// LS Electric XG5000 project: 1조_2차_2축_공압+로드셀_최종
// PLC LSPLC
// module base 0 slot 0: Input/Output Module:XBM-DN/DP32H2 (DC 24V Input/TR Output, 32 points)
// module base 0 slot 1: Internal Positioning:XBF-PO02E (Open Collector Type, 2 Axis)
// module base 0 slot 2: Positioning Module:XBF-PN04B (Position Control, EtherCAT Network Type(4 axis))
// module base 0 slot 3: Loadcell Input Module:XBF-LD02S (Isolated-type Loadcell Input(2 Channels))
// task INIT: Kind=1 Priority=2

PROGRAM ERROR (task: 스캔 프로그램)

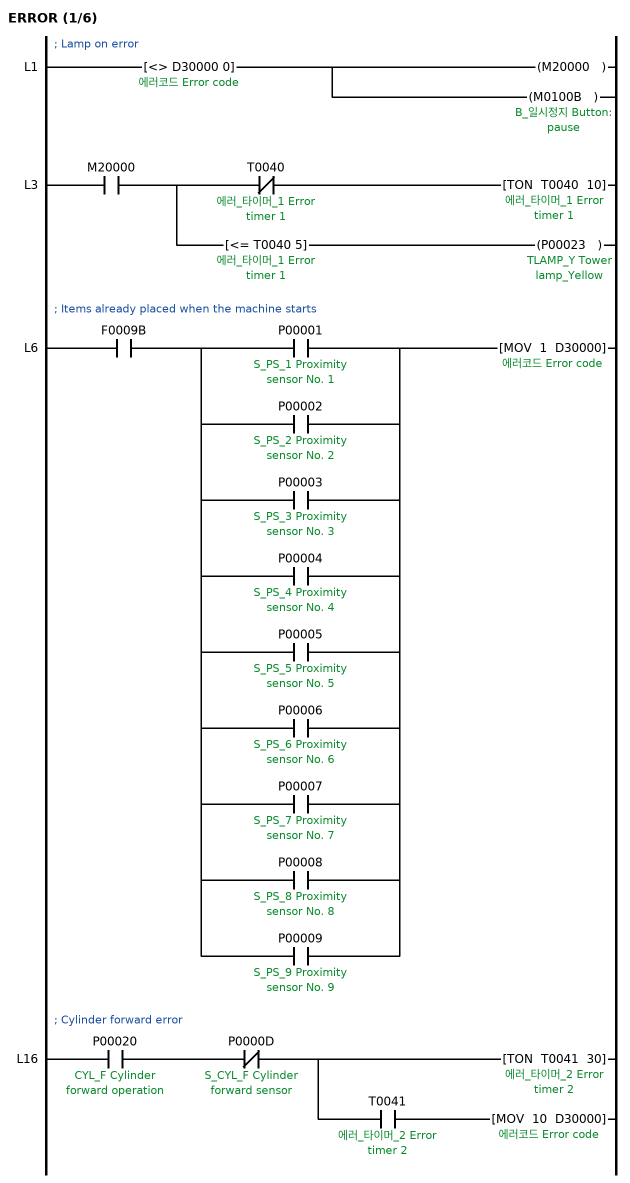
// Lamp on error
; L1
LOAD<>    D30000 0	// 에러코드 Error code
OUT       M20000
OUT       M0100B	// B_일시정지 Button: pause
; L3
LOAD      M20000
MPUSH
AND NOT   T0040	// 에러_타이머_1 Error timer 1
TON       T0040 10	// 에러_타이머_1 Error timer 1
MPOP
AND<=     T0040 5	// 에러_타이머_1 Error timer 1
OUT       P00023	// TLAMP_Y Tower lamp_Yellow
// Items already placed when the machine starts
; L6
LOAD      F0009B
LOAD      P00001	// S_PS_1 Proximity sensor No. 1
OR        P00002	// S_PS_2 Proximity sensor No. 2
OR        P00003	// S_PS_3 Proximity sensor No. 3
OR        P00004	// S_PS_4 Proximity sensor No. 4
OR        P00005	// S_PS_5 Proximity sensor No. 5
OR        P00006	// S_PS_6 Proximity sensor No. 6
OR        P00007	// S_PS_7 Proximity sensor No. 7
OR        P00008	// S_PS_8 Proximity sensor No. 8
OR        P00009	// S_PS_9 Proximity sensor No. 9
AND LOAD
MOV       1 D30000	// 에러코드 Error code
// Cylinder forward error
; L16
LOAD      P00020	// CYL_F Cylinder forward operation
AND NOT   P0000D	// S_CYL_F Cylinder forward sensor
TON       T0041 30	// 에러_타이머_2 Error timer 2
AND       T0041	// 에러_타이머_2 Error timer 2
MOV       10 D30000	// 에러코드 Error code

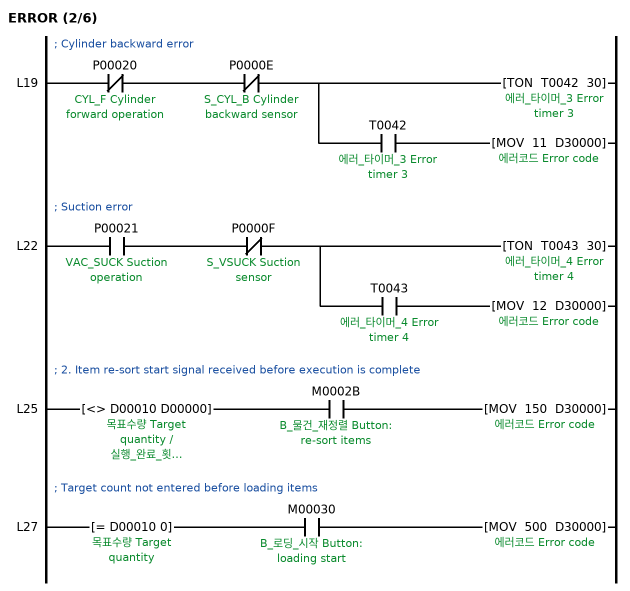
// Cylinder backward error
; L19
LOAD NOT  P00020	// CYL_F Cylinder forward operation
AND NOT   P0000E	// S_CYL_B Cylinder backward sensor
TON       T0042 30	// 에러_타이머_3 Error timer 3
AND       T0042	// 에러_타이머_3 Error timer 3
MOV       11 D30000	// 에러코드 Error code
// Suction error
; L22
LOAD      P00021	// VAC_SUCK Suction operation
AND NOT   P0000F	// S_VSUCK Suction sensor
TON       T0043 30	// 에러_타이머_4 Error timer 4
AND       T0043	// 에러_타이머_4 Error timer 4
MOV       12 D30000	// 에러코드 Error code
// 2. Item re-sort start signal received before execution is complete
; L25
LOAD<>    D00010 D00000	// 목표수량 Target quantity / 실행_완료_횟수 Execution complete count
AND       M0002B	// B_물건_재정렬 Button: re-sort items
MOV       150 D30000	// 에러코드 Error code
// Target count not entered before loading items
; L27
LOAD=     D00010 0	// 목표수량 Target quantity
AND       M00030	// B_로딩_시작 Button: loading start
MOV       500 D30000	// 에러코드 Error code

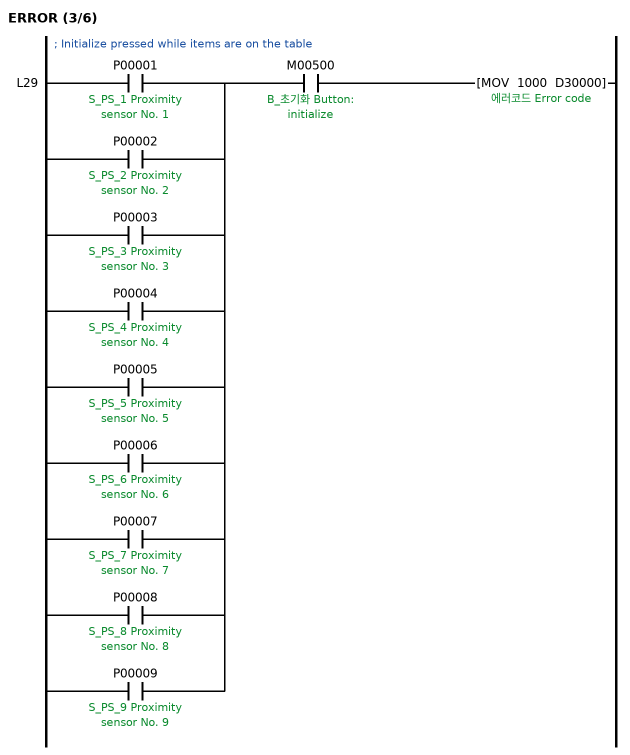
// Initialize pressed while items are on the table
; L29
LOAD      P00001	// S_PS_1 Proximity sensor No. 1
OR        P00002	// S_PS_2 Proximity sensor No. 2
OR        P00003	// S_PS_3 Proximity sensor No. 3
OR        P00004	// S_PS_4 Proximity sensor No. 4
OR        P00005	// S_PS_5 Proximity sensor No. 5
OR        P00006	// S_PS_6 Proximity sensor No. 6
OR        P00007	// S_PS_7 Proximity sensor No. 7
OR        P00008	// S_PS_8 Proximity sensor No. 8
OR        P00009	// S_PS_9 Proximity sensor No. 9
AND       M00500	// B_초기화 Button: initialize
MOV       1000 D30000	// 에러코드 Error code

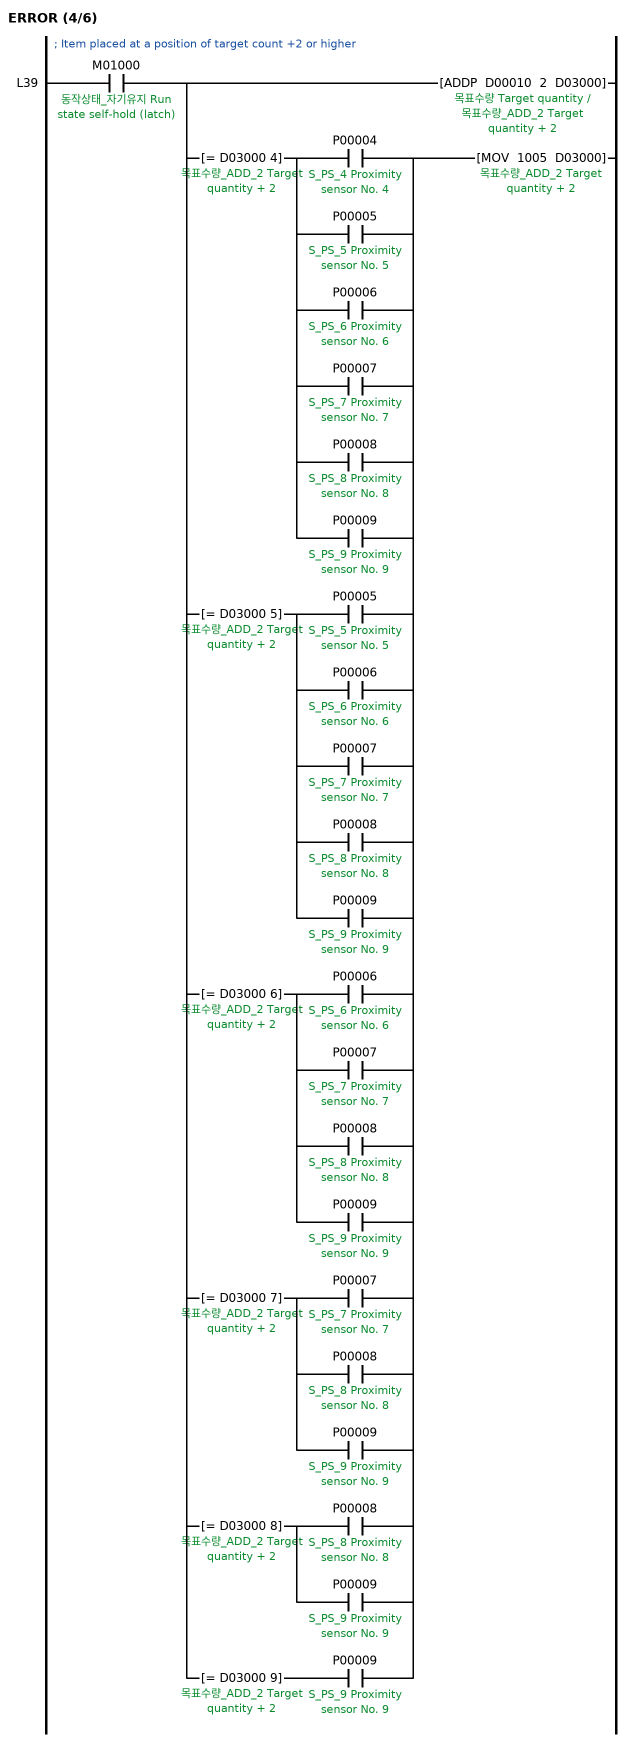
// Item placed at a position of target count +2 or higher
; L39
LOAD      M01000	// 동작상태_자기유지 Run state self-hold (latch)
ADDP      D00010 2 D03000	// 목표수량 Target quantity / 목표수량_ADD_2 Target quantity + 2
LOAD=     D03000 4	// 목표수량_ADD_2 Target quantity + 2
LOAD      P00004	// S_PS_4 Proximity sensor No. 4
OR        P00005	// S_PS_5 Proximity sensor No. 5
OR        P00006	// S_PS_6 Proximity sensor No. 6
OR        P00007	// S_PS_7 Proximity sensor No. 7
OR        P00008	// S_PS_8 Proximity sensor No. 8
OR        P00009	// S_PS_9 Proximity sensor No. 9
AND LOAD
LOAD=     D03000 5	// 목표수량_ADD_2 Target quantity + 2
LOAD      P00005	// S_PS_5 Proximity sensor No. 5
OR        P00006	// S_PS_6 Proximity sensor No. 6
OR        P00007	// S_PS_7 Proximity sensor No. 7
OR        P00008	// S_PS_8 Proximity sensor No. 8
OR        P00009	// S_PS_9 Proximity sensor No. 9
AND LOAD
OR LOAD
LOAD=     D03000 6	// 목표수량_ADD_2 Target quantity + 2
LOAD      P00006	// S_PS_6 Proximity sensor No. 6
OR        P00007	// S_PS_7 Proximity sensor No. 7
OR        P00008	// S_PS_8 Proximity sensor No. 8
OR        P00009	// S_PS_9 Proximity sensor No. 9
AND LOAD
OR LOAD
LOAD=     D03000 7	// 목표수량_ADD_2 Target quantity + 2
LOAD      P00007	// S_PS_7 Proximity sensor No. 7
OR        P00008	// S_PS_8 Proximity sensor No. 8
OR        P00009	// S_PS_9 Proximity sensor No. 9
AND LOAD
OR LOAD
LOAD=     D03000 8	// 목표수량_ADD_2 Target quantity + 2
LOAD      P00008	// S_PS_8 Proximity sensor No. 8
OR        P00009	// S_PS_9 Proximity sensor No. 9
AND LOAD
OR LOAD
LOAD=     D03000 9	// 목표수량_ADD_2 Target quantity + 2
AND       P00009	// S_PS_9 Proximity sensor No. 9
OR LOAD
AND LOAD
MOV       1005 D03000	// 목표수량_ADD_2 Target quantity + 2

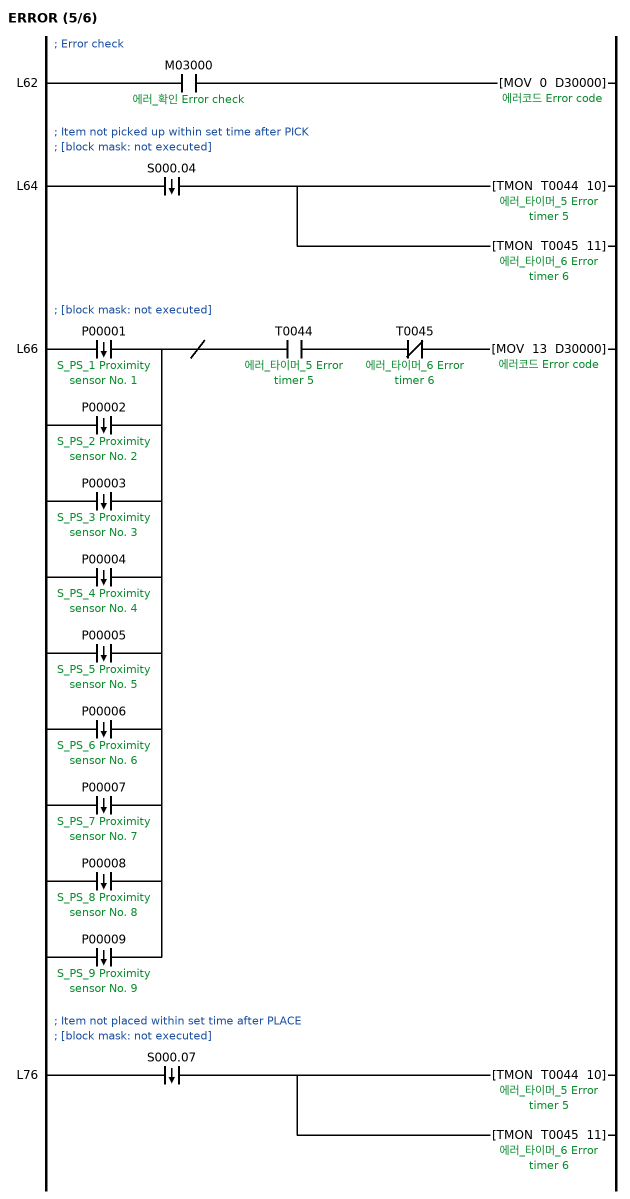
// Error check
; L62
LOAD      M03000	// 에러_확인 Error check
MOV       0 D30000	// 에러코드 Error code
// Item not picked up within set time after PICK
; L64 (block mask: not executed)
LOADN     S000.04
TMON      T0044 10	// 에러_타이머_5 Error timer 5
TMON      T0045 11	// 에러_타이머_6 Error timer 6
; L66 (block mask: not executed)
LOADN     P00001	// S_PS_1 Proximity sensor No. 1
ORN       P00002	// S_PS_2 Proximity sensor No. 2
ORN       P00003	// S_PS_3 Proximity sensor No. 3
ORN       P00004	// S_PS_4 Proximity sensor No. 4
ORN       P00005	// S_PS_5 Proximity sensor No. 5
ORN       P00006	// S_PS_6 Proximity sensor No. 6
ORN       P00007	// S_PS_7 Proximity sensor No. 7
ORN       P00008	// S_PS_8 Proximity sensor No. 8
ORN       P00009	// S_PS_9 Proximity sensor No. 9
NOT
AND       T0044	// 에러_타이머_5 Error timer 5
AND NOT   T0045	// 에러_타이머_6 Error timer 6
MOV       13 D30000	// 에러코드 Error code
// Item not placed within set time after PLACE
; L76 (block mask: not executed)
LOADN     S000.07
TMON      T0044 10	// 에러_타이머_5 Error timer 5
TMON      T0045 11	// 에러_타이머_6 Error timer 6

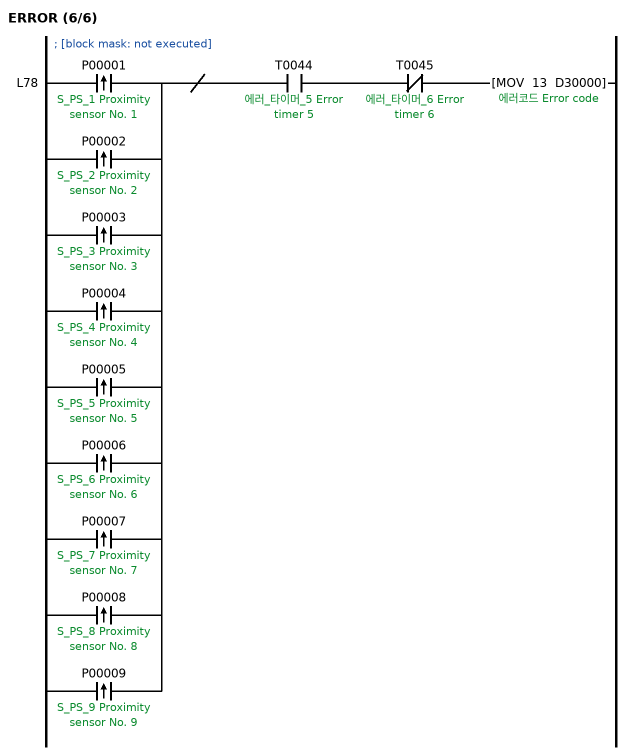
; L78 (block mask: not executed)
LOADP     P00001	// S_PS_1 Proximity sensor No. 1
ORP       P00002	// S_PS_2 Proximity sensor No. 2
ORP       P00003	// S_PS_3 Proximity sensor No. 3
ORP       P00004	// S_PS_4 Proximity sensor No. 4
ORP       P00005	// S_PS_5 Proximity sensor No. 5
ORP       P00006	// S_PS_6 Proximity sensor No. 6
ORP       P00007	// S_PS_7 Proximity sensor No. 7
ORP       P00008	// S_PS_8 Proximity sensor No. 8
ORP       P00009	// S_PS_9 Proximity sensor No. 9
NOT
AND       T0044	// 에러_타이머_5 Error timer 5
AND NOT   T0045	// 에러_타이머_6 Error timer 6
MOV       13 D30000	// 에러코드 Error code

PROGRAM Servo (task: 스캔 프로그램)

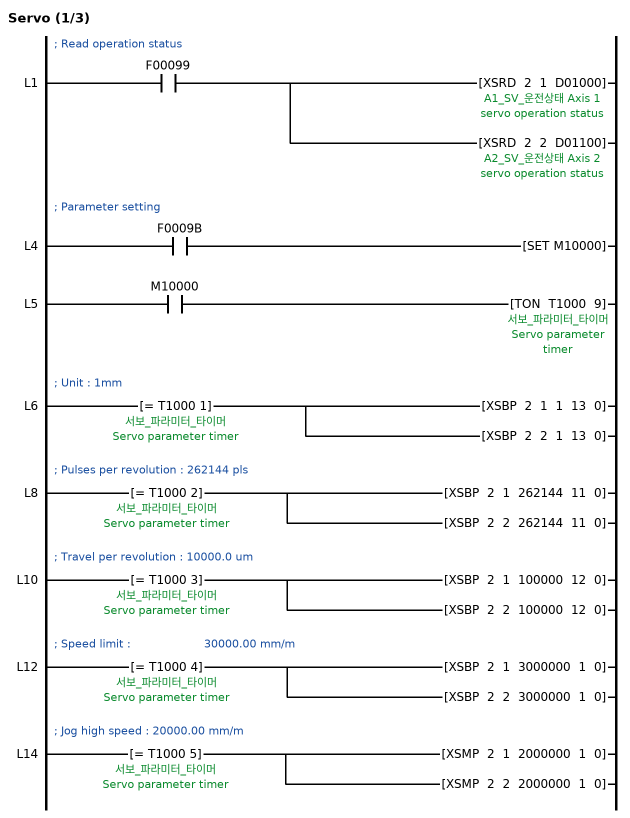
// Read operation status
; L1
LOAD      F00099
XSRD      2 1 D01000	// A1_SV_운전상태 Axis 1 servo operation status
XSRD      2 2 D01100	// A2_SV_운전상태 Axis 2 servo operation status
// Parameter setting
; L4
LOAD      F0009B
SET       M10000
; L5
LOAD      M10000
TON       T1000 9	// 서보_파라미터_타이머 Servo parameter timer
; L6
LOAD=     T1000 1	// 서보_파라미터_타이머 Servo parameter timer
XSBP      2 1 1 13 0
XSBP      2 2 1 13 0
// output comment: Unit : 1mm
; L8
LOAD=     T1000 2	// 서보_파라미터_타이머 Servo parameter timer
XSBP      2 1 262144 11 0
XSBP      2 2 262144 11 0
// output comment: Pulses per revolution : 262144 pls
; L10
LOAD=     T1000 3	// 서보_파라미터_타이머 Servo parameter timer
XSBP      2 1 100000 12 0
XSBP      2 2 100000 12 0
// output comment: Travel per revolution : 10000.0 um
; L12
LOAD=     T1000 4	// 서보_파라미터_타이머 Servo parameter timer
XSBP      2 1 3000000 1 0
XSBP      2 2 3000000 1 0
// output comment: Speed limit :                     30000.00 mm/m
; L14
LOAD=     T1000 5	// 서보_파라미터_타이머 Servo parameter timer
XSMP      2 1 2000000 1 0
XSMP      2 2 2000000 1 0
// output comment: Jog high speed : 20000.00 mm/m

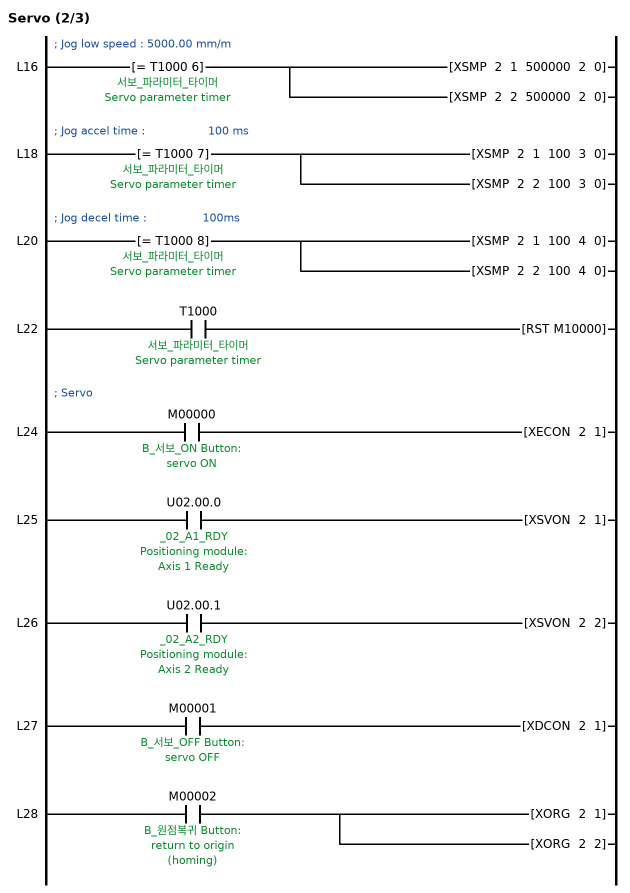
; L16
LOAD=     T1000 6	// 서보_파라미터_타이머 Servo parameter timer
XSMP      2 1 500000 2 0
XSMP      2 2 500000 2 0
// output comment: Jog low speed : 5000.00 mm/m
; L18
LOAD=     T1000 7	// 서보_파라미터_타이머 Servo parameter timer
XSMP      2 1 100 3 0
XSMP      2 2 100 3 0
// output comment: Jog accel time :                  100 ms
; L20
LOAD=     T1000 8	// 서보_파라미터_타이머 Servo parameter timer
XSMP      2 1 100 4 0
XSMP      2 2 100 4 0
// output comment: Jog decel time :                100ms
; L22
LOAD      T1000	// 서보_파라미터_타이머 Servo parameter timer
RST       M10000
// Servo
; L24
LOAD      M00000	// B_서보_ON Button: servo ON
XECON     2 1
; L25
LOAD      U02.00.0	// _02_A1_RDY Positioning module: Axis 1 Ready
XSVON     2 1
; L26
LOAD      U02.00.1	// _02_A2_RDY Positioning module: Axis 2 Ready
XSVON     2 2
; L27
LOAD      M00001	// B_서보_OFF Button: servo OFF
XDCON     2 1
; L28
LOAD      M00002	// B_원점복귀 Button: return to origin (homing)
XORG      2 1
XORG      2 2

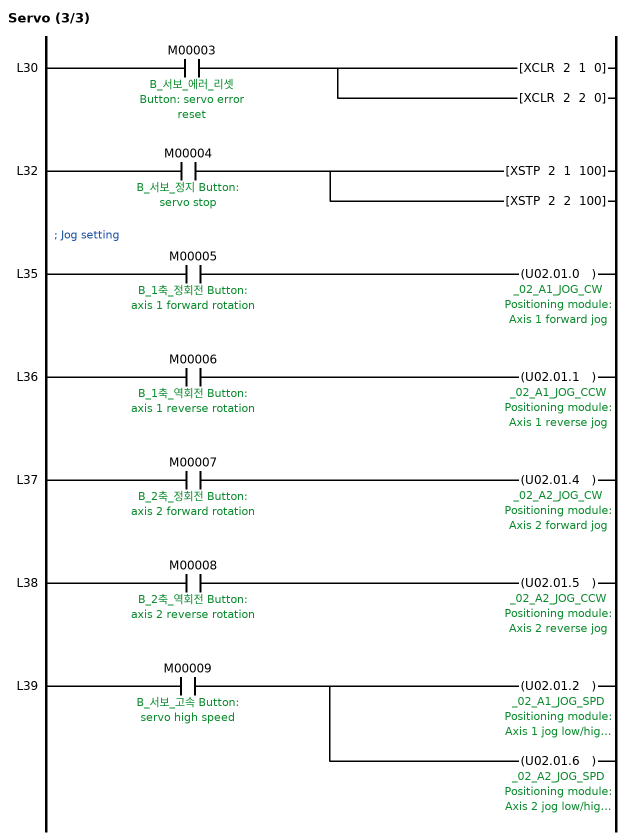
; L30
LOAD      M00003	// B_서보_에러_리셋 Button: servo error reset
XCLR      2 1 0
XCLR      2 2 0
; L32
LOAD      M00004	// B_서보_정지 Button: servo stop
XSTP      2 1 100
XSTP      2 2 100
// Jog setting
; L35
LOAD      M00005	// B_1축_정회전 Button: axis 1 forward rotation
OUT       U02.01.0	// _02_A1_JOG_CW Positioning module: Axis 1 forward jog
; L36
LOAD      M00006	// B_1축_역회전 Button: axis 1 reverse rotation
OUT       U02.01.1	// _02_A1_JOG_CCW Positioning module: Axis 1 reverse jog
; L37
LOAD      M00007	// B_2축_정회전 Button: axis 2 forward rotation
OUT       U02.01.4	// _02_A2_JOG_CW Positioning module: Axis 2 forward jog
; L38
LOAD      M00008	// B_2축_역회전 Button: axis 2 reverse rotation
OUT       U02.01.5	// _02_A2_JOG_CCW Positioning module: Axis 2 reverse jog
; L39
LOAD      M00009	// B_서보_고속 Button: servo high speed
OUT       U02.01.2	// _02_A1_JOG_SPD Positioning module: Axis 1 jog low/high speed
OUT       U02.01.6	// _02_A2_JOG_SPD Positioning module: Axis 2 jog low/high speed

PROGRAM Load_Cell (task: 스캔 프로그램)

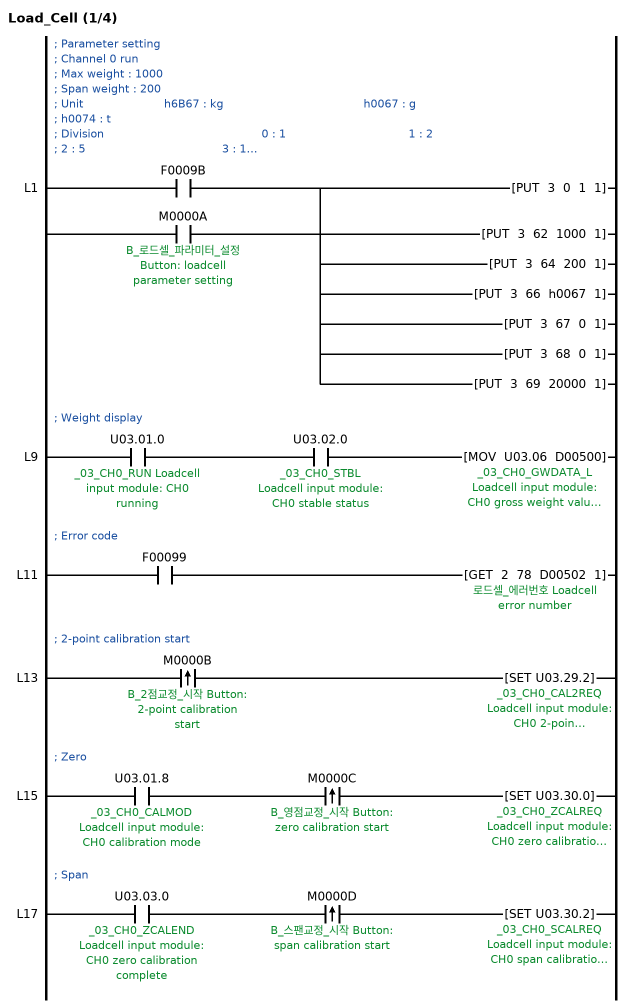
// Parameter setting
; L1
LOAD      F0009B
OR        M0000A	// B_로드셀_파라미터_설정 Button: loadcell parameter setting
PUT       3 0 1 1
PUT       3 62 1000 1
PUT       3 64 200 1
PUT       3 66 h0067 1
PUT       3 67 0 1
PUT       3 68 0 1
PUT       3 69 20000 1
// output comment: Channel 0 run
// output comment: Max weight : 1000
// output comment: Span weight : 200
// output comment: Unit                       h6B67 : kg                                        h0067 : g                                         h0074 : t
// output comment: Division                                             0 : 1                                   1 : 2                                             2 : 5                                       3 : 10
// output comment: Decimal                    0 : 1                    1: 0.1                         2 : 0.01                  3 : 0.001
// output comment: Loadcell sensitivity : 2mV/V
// Weight display
; L9
LOAD      U03.01.0	// _03_CH0_RUN Loadcell input module: CH0 running
AND       U03.02.0	// _03_CH0_STBL Loadcell input module: CH0 stable status
MOV       U03.06 D00500	// _03_CH0_GWDATA_L Loadcell input module: CH0 gross weight value (low) / Mass
// Error code
; L11
LOAD      F00099
GET       2 78 D00502 1	// 로드셀_에러번호 Loadcell error number
// 2-point calibration start
; L13
LOADP     M0000B	// B_2점교정_시작 Button: 2-point calibration start
SET       U03.29.2	// _03_CH0_CAL2REQ Loadcell input module: CH0 2-point calibration mode request
// Zero
; L15
LOAD      U03.01.8	// _03_CH0_CALMOD Loadcell input module: CH0 calibration mode
ANDP      M0000C	// B_영점교정_시작 Button: zero calibration start
SET       U03.30.0	// _03_CH0_ZCALREQ Loadcell input module: CH0 zero calibration command
// Span
; L17
LOAD      U03.03.0	// _03_CH0_ZCALEND Loadcell input module: CH0 zero calibration complete
ANDP      M0000D	// B_스팬교정_시작 Button: span calibration start
SET       U03.30.2	// _03_CH0_SCALREQ Loadcell input module: CH0 span calibration command

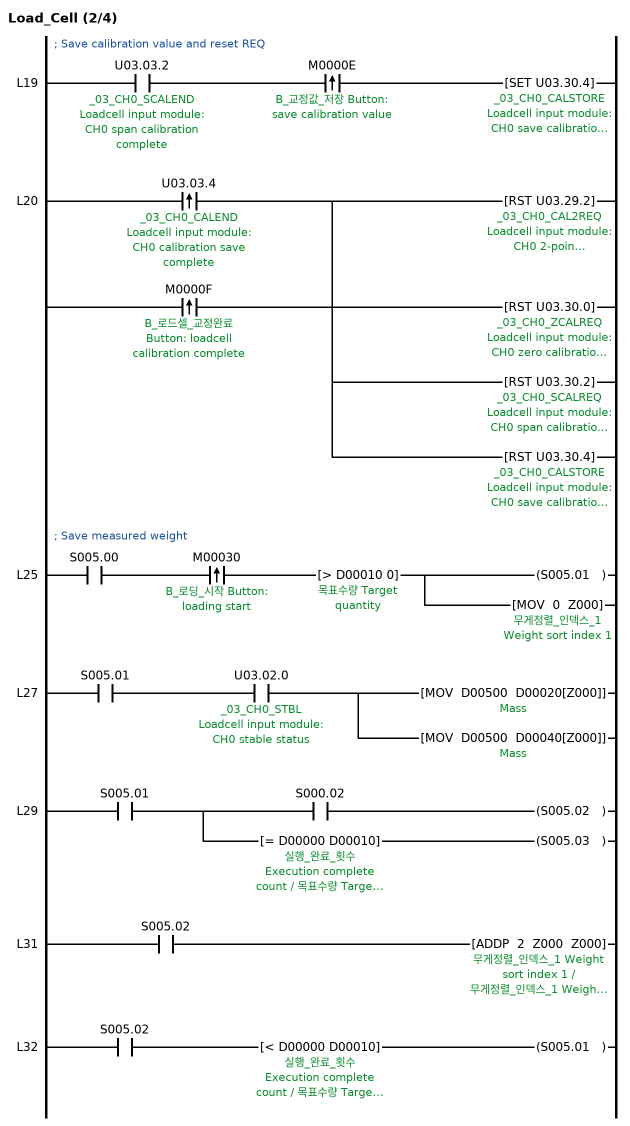
// Save calibration value and reset REQ
; L19
LOAD      U03.03.2	// _03_CH0_SCALEND Loadcell input module: CH0 span calibration complete
ANDP      M0000E	// B_교정값_저장 Button: save calibration value
SET       U03.30.4	// _03_CH0_CALSTORE Loadcell input module: CH0 save calibration value command
; L20
LOADP     U03.03.4	// _03_CH0_CALEND Loadcell input module: CH0 calibration save complete
ORP       M0000F	// B_로드셀_교정완료 Button: loadcell calibration complete
RST       U03.29.2	// _03_CH0_CAL2REQ Loadcell input module: CH0 2-point calibration mode request
RST       U03.30.0	// _03_CH0_ZCALREQ Loadcell input module: CH0 zero calibration command
RST       U03.30.2	// _03_CH0_SCALREQ Loadcell input module: CH0 span calibration command
RST       U03.30.4	// _03_CH0_CALSTORE Loadcell input module: CH0 save calibration value command
// Save measured weight
; L25
LOAD      S005.00
ANDP      M00030	// B_로딩_시작 Button: loading start
AND>      D00010 0	// 목표수량 Target quantity
OUT       S005.01
MOV       0 Z000	// 무게정렬_인덱스_1 Weight sort index 1
; L27
LOAD      S005.01
AND       U03.02.0	// _03_CH0_STBL Loadcell input module: CH0 stable status
MOV       D00500 D00020[Z000]	// Mass
MOV       D00500 D00040[Z000]	// Mass
; L29
LOAD      S005.01
MPUSH
AND       S000.02
OUT       S005.02
MPOP
AND=      D00000 D00010	// 실행_완료_횟수 Execution complete count / 목표수량 Target quantity
OUT       S005.03
; L31
LOAD      S005.02
ADDP      2 Z000 Z000	// 무게정렬_인덱스_1 Weight sort index 1 / 무게정렬_인덱스_1 Weight sort index 1
; L32
LOAD      S005.02
AND<      D00000 D00010	// 실행_완료_횟수 Execution complete count / 목표수량 Target quantity
OUT       S005.01

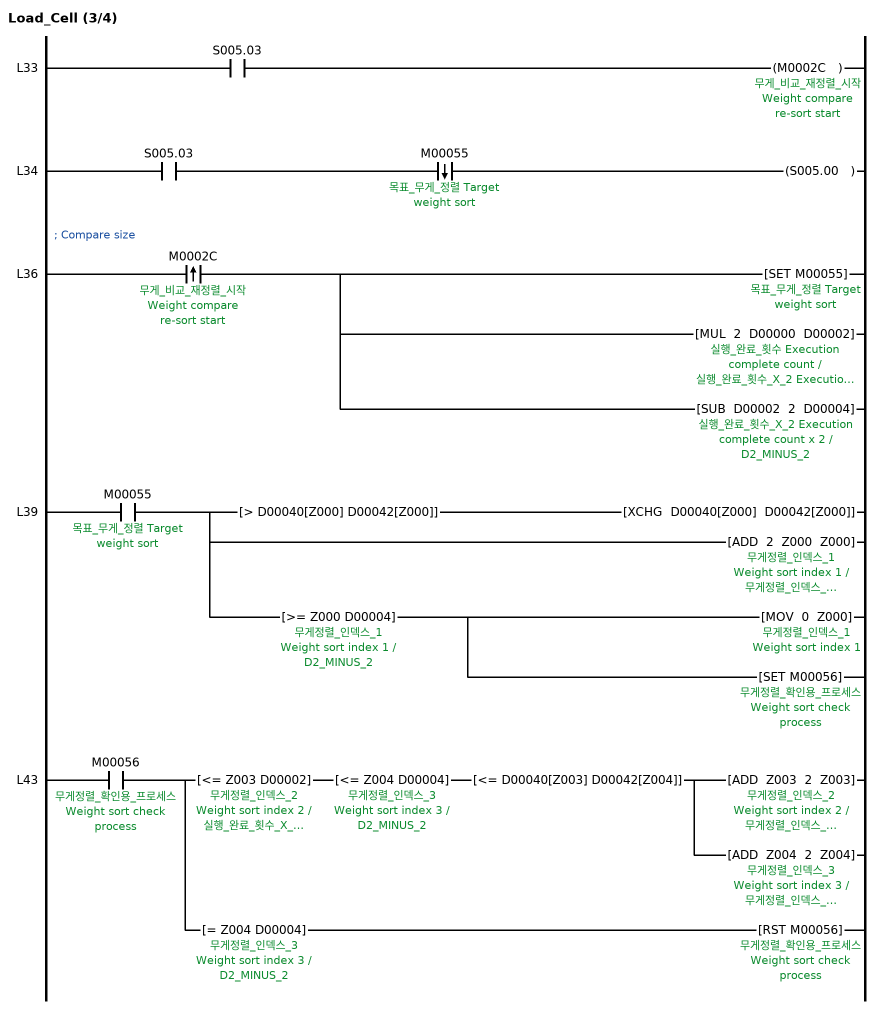
; L33
LOAD      S005.03
OUT       M0002C	// 무게_비교_재정렬_시작 Weight compare re-sort start
; L34
LOAD      S005.03
ANDN      M00055	// 목표_무게_정렬 Target weight sort
OUT       S005.00
// Compare size
; L36
LOADP     M0002C	// 무게_비교_재정렬_시작 Weight compare re-sort start
SET       M00055	// 목표_무게_정렬 Target weight sort
MUL       2 D00000 D00002	// 실행_완료_횟수 Execution complete count / 실행_완료_횟수_X_2 Execution complete count x 2
SUB       D00002 2 D00004	// 실행_완료_횟수_X_2 Execution complete count x 2 / D2_MINUS_2
; L39
LOAD      M00055	// 목표_무게_정렬 Target weight sort
MPUSH
AND>      D00040[Z000] D00042[Z000]
XCHG      D00040[Z000] D00042[Z000]
MPOP
ADD       2 Z000 Z000	// 무게정렬_인덱스_1 Weight sort index 1 / 무게정렬_인덱스_1 Weight sort index 1
AND>=     Z000 D00004	// 무게정렬_인덱스_1 Weight sort index 1 / D2_MINUS_2
MOV       0 Z000	// 무게정렬_인덱스_1 Weight sort index 1
SET       M00056	// 무게정렬_확인용_프로세스 Weight sort check process
; L43
LOAD      M00056	// 무게정렬_확인용_프로세스 Weight sort check process
MPUSH
AND<=     Z003 D00002	// 무게정렬_인덱스_2 Weight sort index 2 / 실행_완료_횟수_X_2 Execution complete count x 2
AND<=     Z004 D00004	// 무게정렬_인덱스_3 Weight sort index 3 / D2_MINUS_2
AND<=     D00040[Z003] D00042[Z004]
ADD       Z003 2 Z003	// 무게정렬_인덱스_2 Weight sort index 2 / 무게정렬_인덱스_2 Weight sort index 2
ADD       Z004 2 Z004	// 무게정렬_인덱스_3 Weight sort index 3 / 무게정렬_인덱스_3 Weight sort index 3
MPOP
AND=      Z004 D00004	// 무게정렬_인덱스_3 Weight sort index 3 / D2_MINUS_2
RST       M00056	// 무게정렬_확인용_프로세스 Weight sort check process

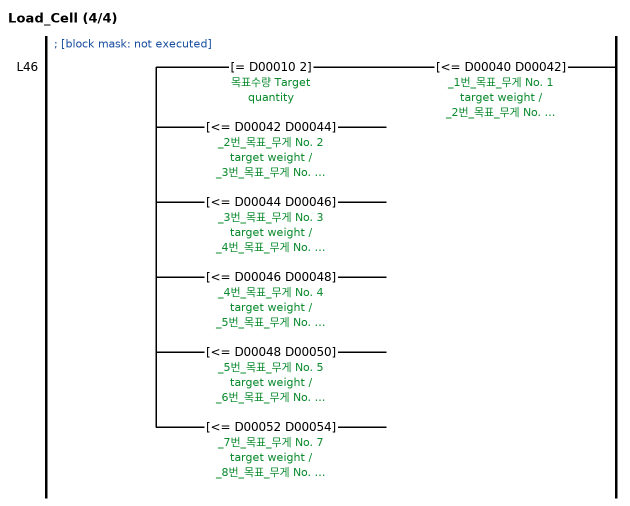
; L46 (block mask: not executed)
// network not rendered as a mnemonic list; see the picture

PROGRAM Pick_&_Place (task: 스캔 프로그램)

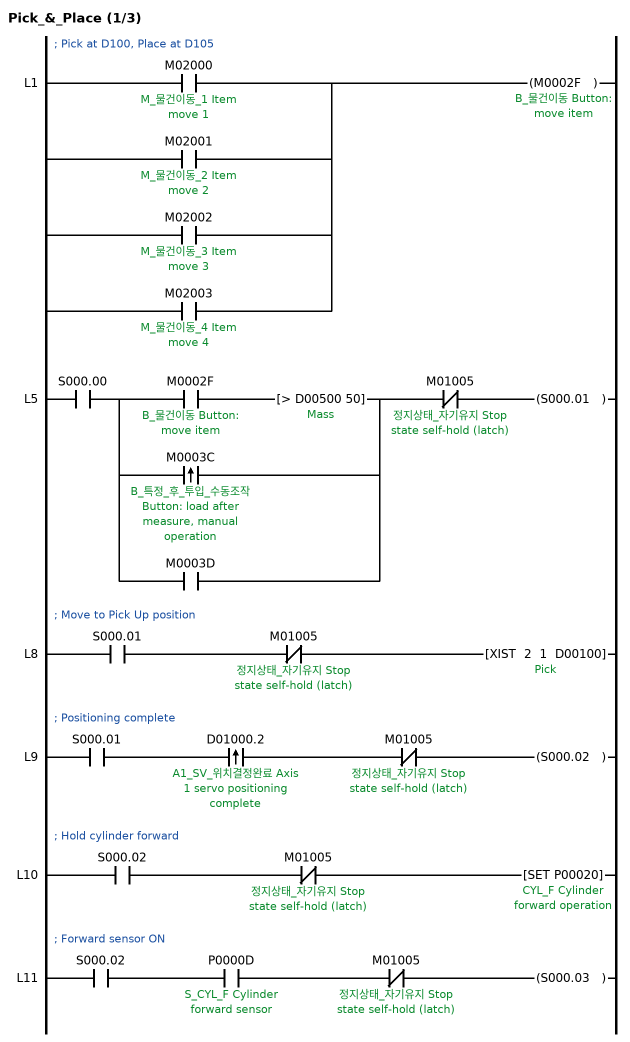
// Pick at D100, Place at D105
; L1
LOAD      M02000	// M_물건이동_1 Item move 1
OR        M02001	// M_물건이동_2 Item move 2
OR        M02002	// M_물건이동_3 Item move 3
OR        M02003	// M_물건이동_4 Item move 4
OUT       M0002F	// B_물건이동 Button: move item
; L5
LOAD      S000.00
LOAD      M0002F	// B_물건이동 Button: move item
AND>      D00500 50	// Mass
ORP       M0003C	// B_특정_후_투입_수동조작 Button: load after measure, manual operation
OR        M0003D
AND LOAD
AND NOT   M01005	// 정지상태_자기유지 Stop state self-hold (latch)
OUT       S000.01
; L8
LOAD      S000.01
AND NOT   M01005	// 정지상태_자기유지 Stop state self-hold (latch)
XIST      2 1 D00100	// Pick
// output comment: Move to Pick Up position
; L9
LOAD      S000.01
ANDP      D01000.2	// A1_SV_위치결정완료 Axis 1 servo positioning complete
AND NOT   M01005	// 정지상태_자기유지 Stop state self-hold (latch)
OUT       S000.02
// output comment: Positioning complete
; L10
LOAD      S000.02
AND NOT   M01005	// 정지상태_자기유지 Stop state self-hold (latch)
SET       P00020	// CYL_F Cylinder forward operation
// output comment: Hold cylinder forward
; L11
LOAD      S000.02
AND       P0000D	// S_CYL_F Cylinder forward sensor
AND NOT   M01005	// 정지상태_자기유지 Stop state self-hold (latch)
OUT       S000.03
// output comment: Forward sensor ON

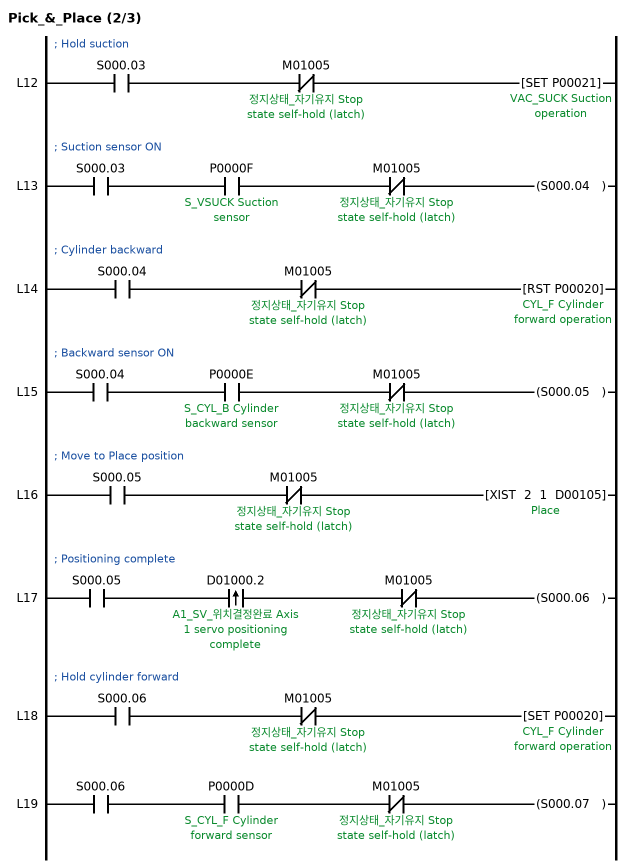
; L12
LOAD      S000.03
AND NOT   M01005	// 정지상태_자기유지 Stop state self-hold (latch)
SET       P00021	// VAC_SUCK Suction operation
// output comment: Hold suction
; L13
LOAD      S000.03
AND       P0000F	// S_VSUCK Suction sensor
AND NOT   M01005	// 정지상태_자기유지 Stop state self-hold (latch)
OUT       S000.04
// output comment: Suction sensor ON
; L14
LOAD      S000.04
AND NOT   M01005	// 정지상태_자기유지 Stop state self-hold (latch)
RST       P00020	// CYL_F Cylinder forward operation
// output comment: Cylinder backward
; L15
LOAD      S000.04
AND       P0000E	// S_CYL_B Cylinder backward sensor
AND NOT   M01005	// 정지상태_자기유지 Stop state self-hold (latch)
OUT       S000.05
// output comment: Backward sensor ON
; L16
LOAD      S000.05
AND NOT   M01005	// 정지상태_자기유지 Stop state self-hold (latch)
XIST      2 1 D00105	// Place
// output comment: Move to Place position
; L17
LOAD      S000.05
ANDP      D01000.2	// A1_SV_위치결정완료 Axis 1 servo positioning complete
AND NOT   M01005	// 정지상태_자기유지 Stop state self-hold (latch)
OUT       S000.06
// output comment: Positioning complete
; L18
LOAD      S000.06
AND NOT   M01005	// 정지상태_자기유지 Stop state self-hold (latch)
SET       P00020	// CYL_F Cylinder forward operation
// output comment: Hold cylinder forward
; L19
LOAD      S000.06
AND       P0000D	// S_CYL_F Cylinder forward sensor
AND NOT   M01005	// 정지상태_자기유지 Stop state self-hold (latch)
OUT       S000.07

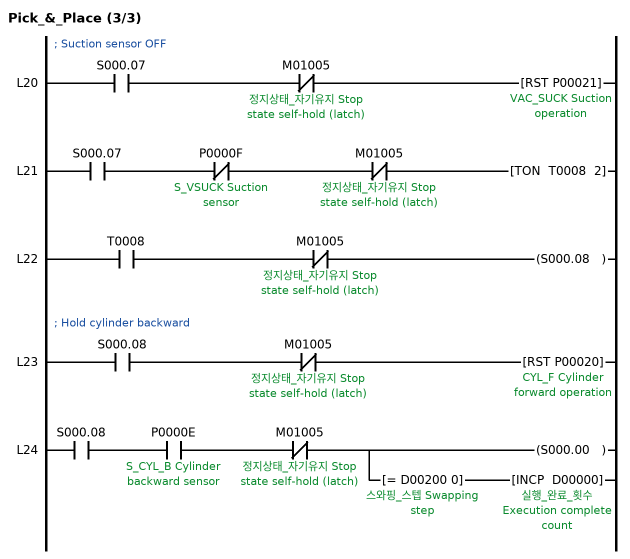
; L20
LOAD      S000.07
AND NOT   M01005	// 정지상태_자기유지 Stop state self-hold (latch)
RST       P00021	// VAC_SUCK Suction operation
// output comment: Suction sensor OFF
; L21
LOAD      S000.07
AND NOT   P0000F	// S_VSUCK Suction sensor
AND NOT   M01005	// 정지상태_자기유지 Stop state self-hold (latch)
TON       T0008 2
; L22
LOAD      T0008
AND NOT   M01005	// 정지상태_자기유지 Stop state self-hold (latch)
OUT       S000.08
; L23
LOAD      S000.08
AND NOT   M01005	// 정지상태_자기유지 Stop state self-hold (latch)
RST       P00020	// CYL_F Cylinder forward operation
// output comment: Hold cylinder backward
; L24
LOAD      S000.08
AND       P0000E	// S_CYL_B Cylinder backward sensor
AND NOT   M01005	// 정지상태_자기유지 Stop state self-hold (latch)
OUT       S000.00
AND=      D00200 0	// 스와핑_스텝 Swapping step
INCP      D00000	// 실행_완료_횟수 Execution complete count

PROGRAM Positioning (task: 스캔 프로그램)

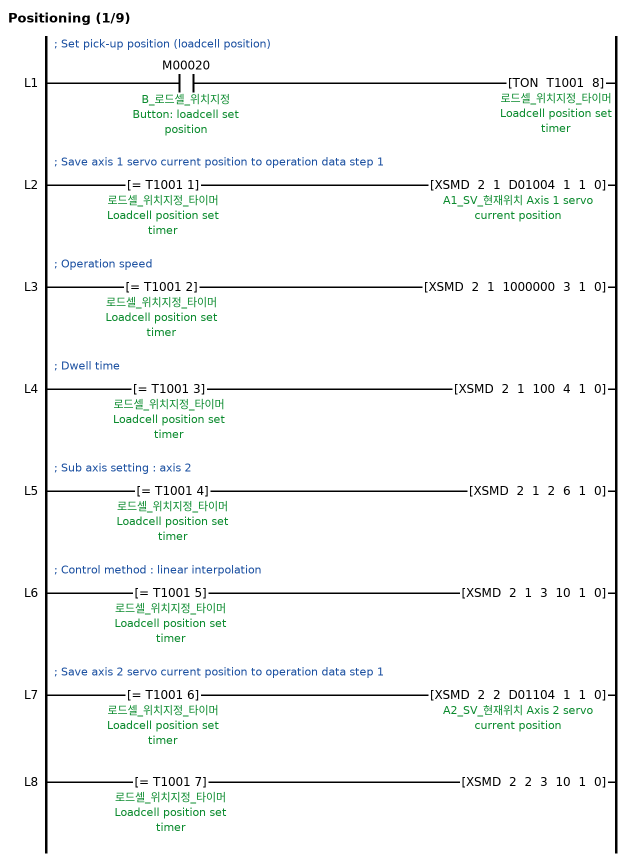
// Set pick-up position (loadcell position)
; L1
LOAD      M00020	// B_로드셀_위치지정 Button: loadcell set position
TON       T1001 8	// 로드셀_위치지정_타이머 Loadcell position set timer
; L2
LOAD=     T1001 1	// 로드셀_위치지정_타이머 Loadcell position set timer
XSMD      2 1 D01004 1 1 0	// A1_SV_현재위치 Axis 1 servo current position
// output comment: Save axis 1 servo current position to operation data step 1
; L3
LOAD=     T1001 2	// 로드셀_위치지정_타이머 Loadcell position set timer
XSMD      2 1 1000000 3 1 0
// output comment: Operation speed
; L4
LOAD=     T1001 3	// 로드셀_위치지정_타이머 Loadcell position set timer
XSMD      2 1 100 4 1 0
// output comment: Dwell time
; L5
LOAD=     T1001 4	// 로드셀_위치지정_타이머 Loadcell position set timer
XSMD      2 1 2 6 1 0
// output comment: Sub axis setting : axis 2
; L6
LOAD=     T1001 5	// 로드셀_위치지정_타이머 Loadcell position set timer
XSMD      2 1 3 10 1 0
// output comment: Control method : linear interpolation
; L7
LOAD=     T1001 6	// 로드셀_위치지정_타이머 Loadcell position set timer
XSMD      2 2 D01104 1 1 0	// A2_SV_현재위치 Axis 2 servo current position
// output comment: Save axis 2 servo current position to operation data step 1
; L8
LOAD=     T1001 7	// 로드셀_위치지정_타이머 Loadcell position set timer
XSMD      2 2 3 10 1 0
// output comment: 

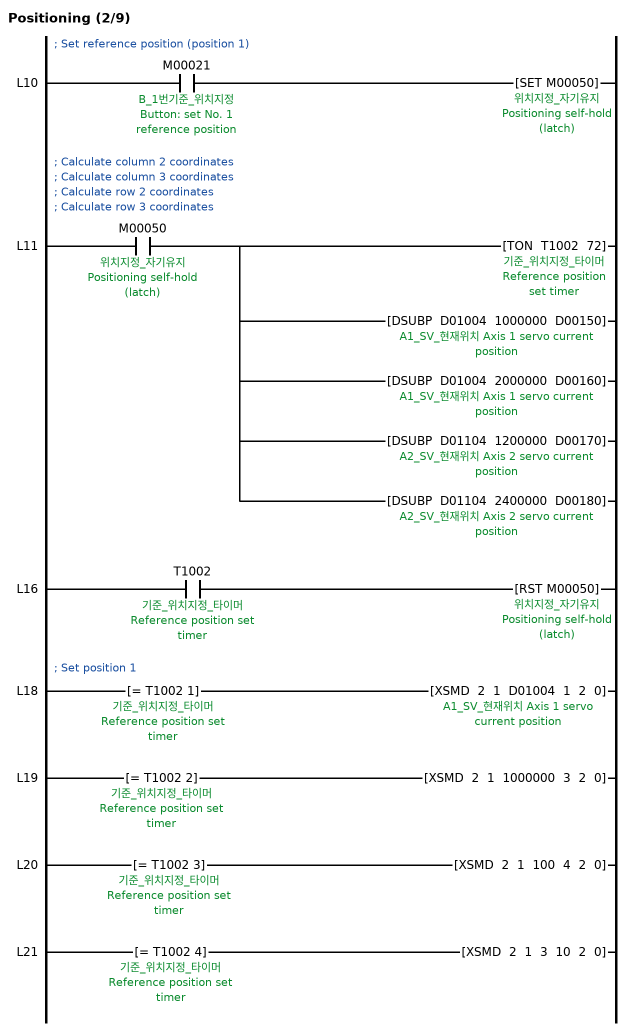
// Set reference position (position 1)
; L10
LOAD      M00021	// B_1번기준_위치지정 Button: set No. 1 reference position
SET       M00050	// 위치지정_자기유지 Positioning self-hold (latch)
; L11
LOAD      M00050	// 위치지정_자기유지 Positioning self-hold (latch)
TON       T1002 72	// 기준_위치지정_타이머 Reference position set timer
DSUBP     D01004 1000000 D00150	// A1_SV_현재위치 Axis 1 servo current position
DSUBP     D01004 2000000 D00160	// A1_SV_현재위치 Axis 1 servo current position
DSUBP     D01104 1200000 D00170	// A2_SV_현재위치 Axis 2 servo current position
DSUBP     D01104 2400000 D00180	// A2_SV_현재위치 Axis 2 servo current position
// output comment: Calculate column 2 coordinates
// output comment: Calculate column 3 coordinates
// output comment: Calculate row 2 coordinates
// output comment: Calculate row 3 coordinates
; L16
LOAD      T1002	// 기준_위치지정_타이머 Reference position set timer
RST       M00050	// 위치지정_자기유지 Positioning self-hold (latch)
// Set position 1
; L18
LOAD=     T1002 1	// 기준_위치지정_타이머 Reference position set timer
XSMD      2 1 D01004 1 2 0	// A1_SV_현재위치 Axis 1 servo current position
; L19
LOAD=     T1002 2	// 기준_위치지정_타이머 Reference position set timer
XSMD      2 1 1000000 3 2 0
; L20
LOAD=     T1002 3	// 기준_위치지정_타이머 Reference position set timer
XSMD      2 1 100 4 2 0
; L21
LOAD=     T1002 4	// 기준_위치지정_타이머 Reference position set timer
XSMD      2 1 3 10 2 0

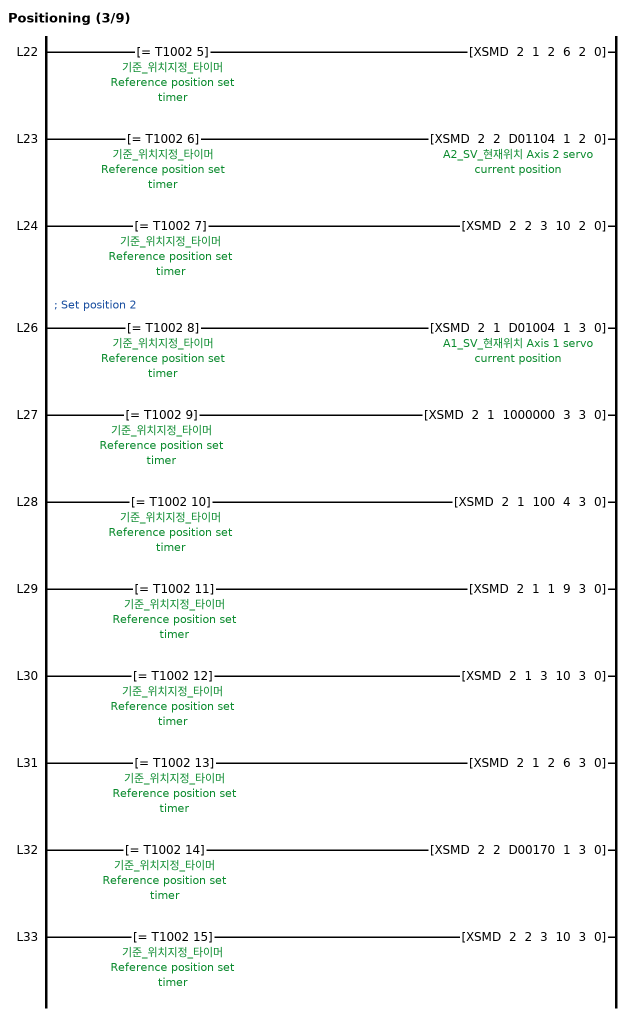
; L22
LOAD=     T1002 5	// 기준_위치지정_타이머 Reference position set timer
XSMD      2 1 2 6 2 0
; L23
LOAD=     T1002 6	// 기준_위치지정_타이머 Reference position set timer
XSMD      2 2 D01104 1 2 0	// A2_SV_현재위치 Axis 2 servo current position
; L24
LOAD=     T1002 7	// 기준_위치지정_타이머 Reference position set timer
XSMD      2 2 3 10 2 0
// Set position 2
; L26
LOAD=     T1002 8	// 기준_위치지정_타이머 Reference position set timer
XSMD      2 1 D01004 1 3 0	// A1_SV_현재위치 Axis 1 servo current position
; L27
LOAD=     T1002 9	// 기준_위치지정_타이머 Reference position set timer
XSMD      2 1 1000000 3 3 0
; L28
LOAD=     T1002 10	// 기준_위치지정_타이머 Reference position set timer
XSMD      2 1 100 4 3 0
; L29
LOAD=     T1002 11	// 기준_위치지정_타이머 Reference position set timer
XSMD      2 1 1 9 3 0
; L30
LOAD=     T1002 12	// 기준_위치지정_타이머 Reference position set timer
XSMD      2 1 3 10 3 0
; L31
LOAD=     T1002 13	// 기준_위치지정_타이머 Reference position set timer
XSMD      2 1 2 6 3 0
; L32
LOAD=     T1002 14	// 기준_위치지정_타이머 Reference position set timer
XSMD      2 2 D00170 1 3 0
; L33
LOAD=     T1002 15	// 기준_위치지정_타이머 Reference position set timer
XSMD      2 2 3 10 3 0

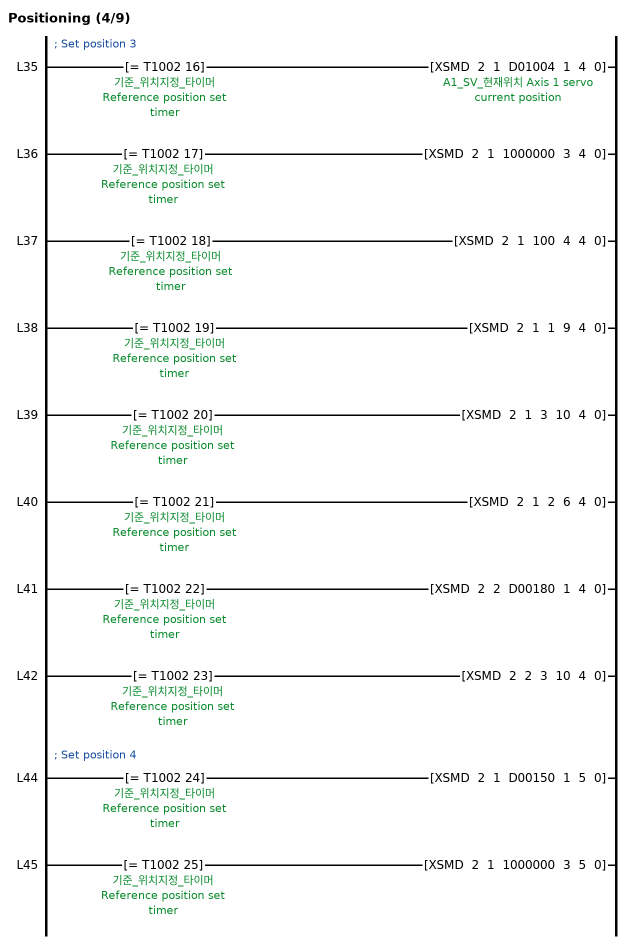
// Set position 3
; L35
LOAD=     T1002 16	// 기준_위치지정_타이머 Reference position set timer
XSMD      2 1 D01004 1 4 0	// A1_SV_현재위치 Axis 1 servo current position
; L36
LOAD=     T1002 17	// 기준_위치지정_타이머 Reference position set timer
XSMD      2 1 1000000 3 4 0
; L37
LOAD=     T1002 18	// 기준_위치지정_타이머 Reference position set timer
XSMD      2 1 100 4 4 0
; L38
LOAD=     T1002 19	// 기준_위치지정_타이머 Reference position set timer
XSMD      2 1 1 9 4 0
; L39
LOAD=     T1002 20	// 기준_위치지정_타이머 Reference position set timer
XSMD      2 1 3 10 4 0
; L40
LOAD=     T1002 21	// 기준_위치지정_타이머 Reference position set timer
XSMD      2 1 2 6 4 0
; L41
LOAD=     T1002 22	// 기준_위치지정_타이머 Reference position set timer
XSMD      2 2 D00180 1 4 0
; L42
LOAD=     T1002 23	// 기준_위치지정_타이머 Reference position set timer
XSMD      2 2 3 10 4 0
// Set position 4
; L44
LOAD=     T1002 24	// 기준_위치지정_타이머 Reference position set timer
XSMD      2 1 D00150 1 5 0
; L45
LOAD=     T1002 25	// 기준_위치지정_타이머 Reference position set timer
XSMD      2 1 1000000 3 5 0

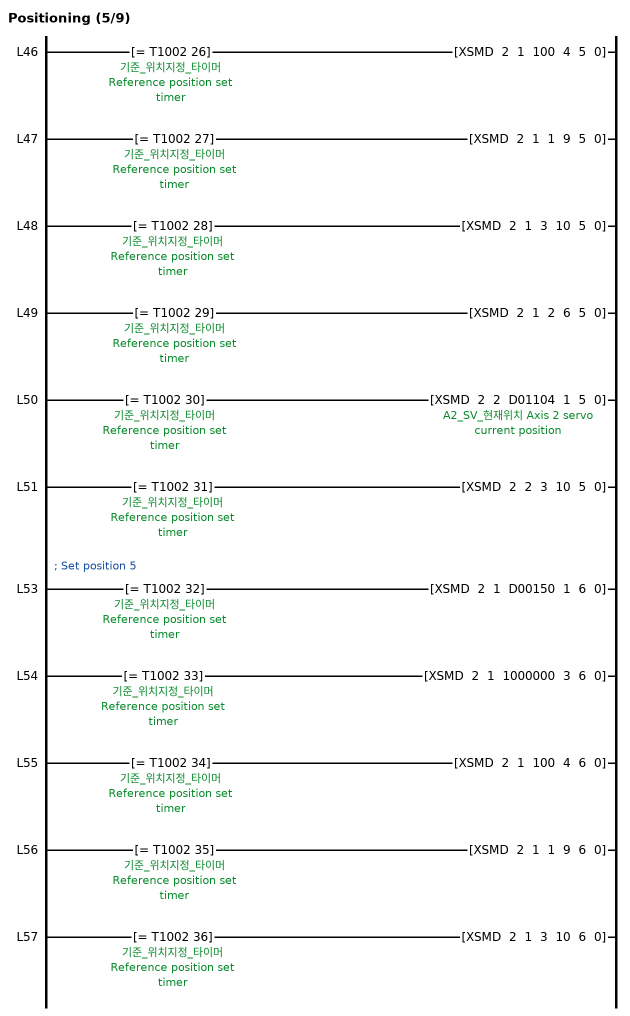
; L46
LOAD=     T1002 26	// 기준_위치지정_타이머 Reference position set timer
XSMD      2 1 100 4 5 0
; L47
LOAD=     T1002 27	// 기준_위치지정_타이머 Reference position set timer
XSMD      2 1 1 9 5 0
; L48
LOAD=     T1002 28	// 기준_위치지정_타이머 Reference position set timer
XSMD      2 1 3 10 5 0
; L49
LOAD=     T1002 29	// 기준_위치지정_타이머 Reference position set timer
XSMD      2 1 2 6 5 0
; L50
LOAD=     T1002 30	// 기준_위치지정_타이머 Reference position set timer
XSMD      2 2 D01104 1 5 0	// A2_SV_현재위치 Axis 2 servo current position
; L51
LOAD=     T1002 31	// 기준_위치지정_타이머 Reference position set timer
XSMD      2 2 3 10 5 0
// Set position 5
; L53
LOAD=     T1002 32	// 기준_위치지정_타이머 Reference position set timer
XSMD      2 1 D00150 1 6 0
; L54
LOAD=     T1002 33	// 기준_위치지정_타이머 Reference position set timer
XSMD      2 1 1000000 3 6 0
; L55
LOAD=     T1002 34	// 기준_위치지정_타이머 Reference position set timer
XSMD      2 1 100 4 6 0
; L56
LOAD=     T1002 35	// 기준_위치지정_타이머 Reference position set timer
XSMD      2 1 1 9 6 0
; L57
LOAD=     T1002 36	// 기준_위치지정_타이머 Reference position set timer
XSMD      2 1 3 10 6 0

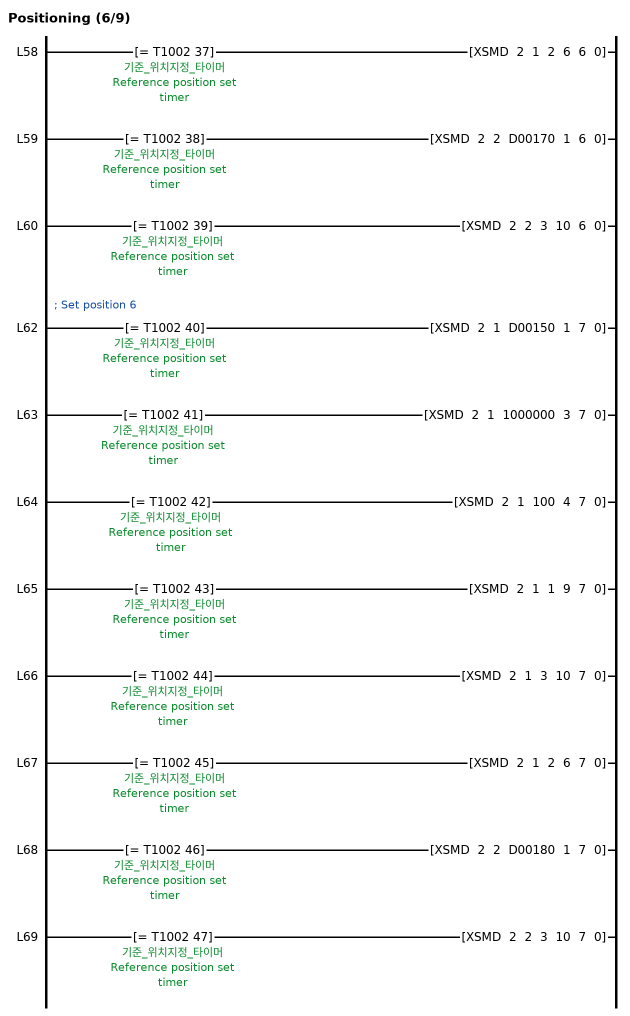
; L58
LOAD=     T1002 37	// 기준_위치지정_타이머 Reference position set timer
XSMD      2 1 2 6 6 0
; L59
LOAD=     T1002 38	// 기준_위치지정_타이머 Reference position set timer
XSMD      2 2 D00170 1 6 0
; L60
LOAD=     T1002 39	// 기준_위치지정_타이머 Reference position set timer
XSMD      2 2 3 10 6 0
// Set position 6
; L62
LOAD=     T1002 40	// 기준_위치지정_타이머 Reference position set timer
XSMD      2 1 D00150 1 7 0
; L63
LOAD=     T1002 41	// 기준_위치지정_타이머 Reference position set timer
XSMD      2 1 1000000 3 7 0
; L64
LOAD=     T1002 42	// 기준_위치지정_타이머 Reference position set timer
XSMD      2 1 100 4 7 0
; L65
LOAD=     T1002 43	// 기준_위치지정_타이머 Reference position set timer
XSMD      2 1 1 9 7 0
; L66
LOAD=     T1002 44	// 기준_위치지정_타이머 Reference position set timer
XSMD      2 1 3 10 7 0
; L67
LOAD=     T1002 45	// 기준_위치지정_타이머 Reference position set timer
XSMD      2 1 2 6 7 0
; L68
LOAD=     T1002 46	// 기준_위치지정_타이머 Reference position set timer
XSMD      2 2 D00180 1 7 0
; L69
LOAD=     T1002 47	// 기준_위치지정_타이머 Reference position set timer
XSMD      2 2 3 10 7 0

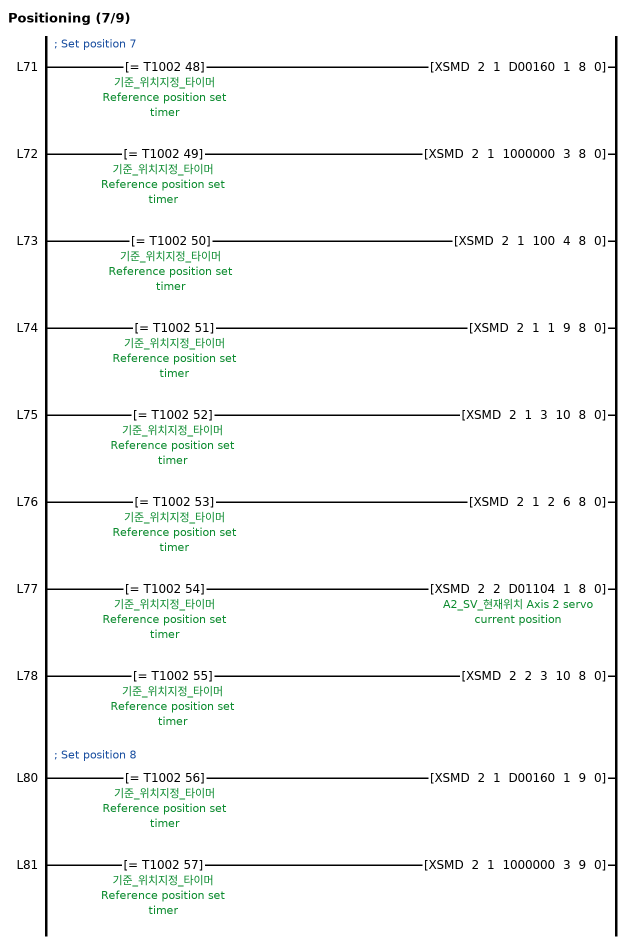
// Set position 7
; L71
LOAD=     T1002 48	// 기준_위치지정_타이머 Reference position set timer
XSMD      2 1 D00160 1 8 0
; L72
LOAD=     T1002 49	// 기준_위치지정_타이머 Reference position set timer
XSMD      2 1 1000000 3 8 0
; L73
LOAD=     T1002 50	// 기준_위치지정_타이머 Reference position set timer
XSMD      2 1 100 4 8 0
; L74
LOAD=     T1002 51	// 기준_위치지정_타이머 Reference position set timer
XSMD      2 1 1 9 8 0
; L75
LOAD=     T1002 52	// 기준_위치지정_타이머 Reference position set timer
XSMD      2 1 3 10 8 0
; L76
LOAD=     T1002 53	// 기준_위치지정_타이머 Reference position set timer
XSMD      2 1 2 6 8 0
; L77
LOAD=     T1002 54	// 기준_위치지정_타이머 Reference position set timer
XSMD      2 2 D01104 1 8 0	// A2_SV_현재위치 Axis 2 servo current position
; L78
LOAD=     T1002 55	// 기준_위치지정_타이머 Reference position set timer
XSMD      2 2 3 10 8 0
// Set position 8
; L80
LOAD=     T1002 56	// 기준_위치지정_타이머 Reference position set timer
XSMD      2 1 D00160 1 9 0
; L81
LOAD=     T1002 57	// 기준_위치지정_타이머 Reference position set timer
XSMD      2 1 1000000 3 9 0

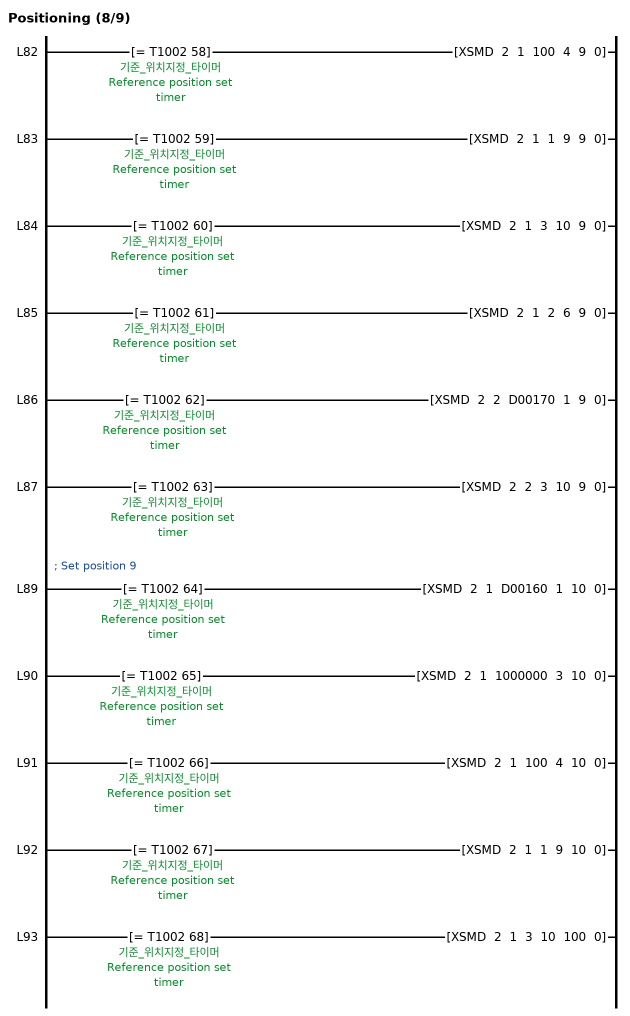
; L82
LOAD=     T1002 58	// 기준_위치지정_타이머 Reference position set timer
XSMD      2 1 100 4 9 0
; L83
LOAD=     T1002 59	// 기준_위치지정_타이머 Reference position set timer
XSMD      2 1 1 9 9 0
; L84
LOAD=     T1002 60	// 기준_위치지정_타이머 Reference position set timer
XSMD      2 1 3 10 9 0
; L85
LOAD=     T1002 61	// 기준_위치지정_타이머 Reference position set timer
XSMD      2 1 2 6 9 0
; L86
LOAD=     T1002 62	// 기준_위치지정_타이머 Reference position set timer
XSMD      2 2 D00170 1 9 0
; L87
LOAD=     T1002 63	// 기준_위치지정_타이머 Reference position set timer
XSMD      2 2 3 10 9 0
// Set position 9
; L89
LOAD=     T1002 64	// 기준_위치지정_타이머 Reference position set timer
XSMD      2 1 D00160 1 10 0
; L90
LOAD=     T1002 65	// 기준_위치지정_타이머 Reference position set timer
XSMD      2 1 1000000 3 10 0
; L91
LOAD=     T1002 66	// 기준_위치지정_타이머 Reference position set timer
XSMD      2 1 100 4 10 0
; L92
LOAD=     T1002 67	// 기준_위치지정_타이머 Reference position set timer
XSMD      2 1 1 9 10 0
; L93
LOAD=     T1002 68	// 기준_위치지정_타이머 Reference position set timer
XSMD      2 1 3 10 100 0

